(* IEC 61131-3 sources: plc-vscode/tests/st/all/trust-platform/examples/OSCAT/conveyor_pulse/non-oop/src, 3 files *)

(* ---- Configuration.st ---- *)
CONFIGURATION ConveyorPulseClassicConfiguration
RESOURCE Cpu0 ON PLC
    TASK MainTask (INTERVAL := T#100ms, PRIORITY := 1);
    PROGRAM Main WITH MainTask : Main;
END_RESOURCE
END_CONFIGURATION

(* ---- Main.st ---- *)
PROGRAM Main
VAR
    BeltPulse : GEN_PULSE;
    ConveyorEnabled : BOOL := FALSE;
    PulseCommand : BOOL;
END_VAR

BeltPulse(ENQ := ConveyorEnabled, PTH := T#500ms, PTL := T#500ms);
PulseCommand := BeltPulse.Q;
END_PROGRAM

(* ---- Tests.st ---- *)
TEST_PROGRAM ConveyorPulseClassicRemainsLowWhenDisabled
VAR
    BeltPulse : GEN_PULSE;
END_VAR

BeltPulse(ENQ := FALSE, PTH := T#500ms, PTL := T#500ms);

ASSERT_FALSE(IN := BeltPulse.Q);
END_TEST_PROGRAM
